# EPICS substitutions: db/Beckhoff_7XXX/ecmcEL7037.substitutions
file "ecmcEL7037-chX.template"
{
  pattern {CH_ID}
          {01   }
}

file "ecmcEL5101-chX.template"
{
  pattern {CH_ID}
          {01   }
}

file "ecmcEL7037_motorLoad-chX.template"
{
  pattern {CH_ID}
          {01   }
}
